SUBAPPLICATION AUF_AB_Softkey_Aux_DataPanel_QXA_SB (* Manuell Auf/Ab mit SoftKey+AUX auf DataPanel-MI-Ausgaenge, Anforderung Sperrblock *)
  (* Standard: 61499-2; Description: Copyright (c) 2026 Meisterschulen am Ostbahnhof This program and the accompanying materials are made available under the terms of the Eclipse Public License 2.0 which is available at https://www.eclipse.org/legal/epl-2.0/ SPDX-License-Identifier: EPL-2.0 *)
  (* Version 1.0, 2026-10-31, Franz Höpfinger, Meisterschulen am Ostbahnhof, Aus Getreidehacke func/Manual/ManFunc_AUF_AB3 in MyLib::sys verschoben und umbenannt, INIT/INITO/QI/QO ergaenzt, u8SAMember als Parameter. *)
  PACKAGE MyLib::sys;
  IMPORT isobus::UT::Q::const::IDs::ID_NULL;
  IMPORT DataPanel::io::MI::DQ::DataPanel_MI_DO_S;
  IMPORT DataPanel::io::MI::DQ::DataPanel_MI_DO;
  IMPORT DataPanel::io::MI::const::MI;
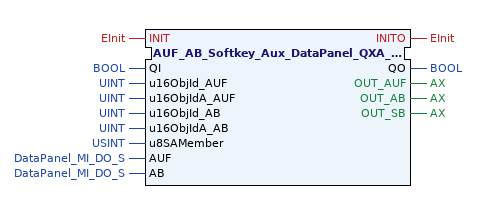
  EVENT_INPUT
    INIT : EInit; (* Initialization Request *)
  END_EVENT
  EVENT_OUTPUT
    INITO : EInit; (* Initialization Confirm *)
  END_EVENT
  VAR_INPUT
    QI : BOOL := TRUE; (* Quality Input - TRUE to enable service *)
    u16ObjId_AUF : UINT := ID_NULL; (* Object ID SoftKey AUF *)
    u16ObjIdA_AUF : UINT := ID_NULL; (* Object ID AuxFunction2 AUF *)
    u16ObjId_AB : UINT := ID_NULL; (* Object ID SoftKey AB *)
    u16ObjIdA_AB : UINT := ID_NULL; (* Object ID AuxFunction2 AB *)
    u8SAMember : USINT := MI::MI_00; (* DataPanel-MI-Modul (Source Address) *)
    AUF : DataPanel::io::MI::DQ::DataPanel_MI_DO_S := DataPanel_MI_DO::Invalid; (* DataPanel-MI-Ausgang AUF *)
    AB : DataPanel::io::MI::DQ::DataPanel_MI_DO_S := DataPanel_MI_DO::Invalid; (* DataPanel-MI-Ausgang AB *)
  END_VAR
  VAR_OUTPUT
    QO : BOOL; (* Quality Output - TRUE if service executed successfully *)
  END_VAR
  PLUGS
    OUT_AUF : adapter::types::unidirectional::AX; (* AUF aktiv *)
    OUT_AB : adapter::types::unidirectional::AX; (* AB aktiv *)
    OUT_SB : adapter::types::unidirectional::AX; (* Sperrblock anfordern (AUF ODER AB) *)
  END_PLUGS
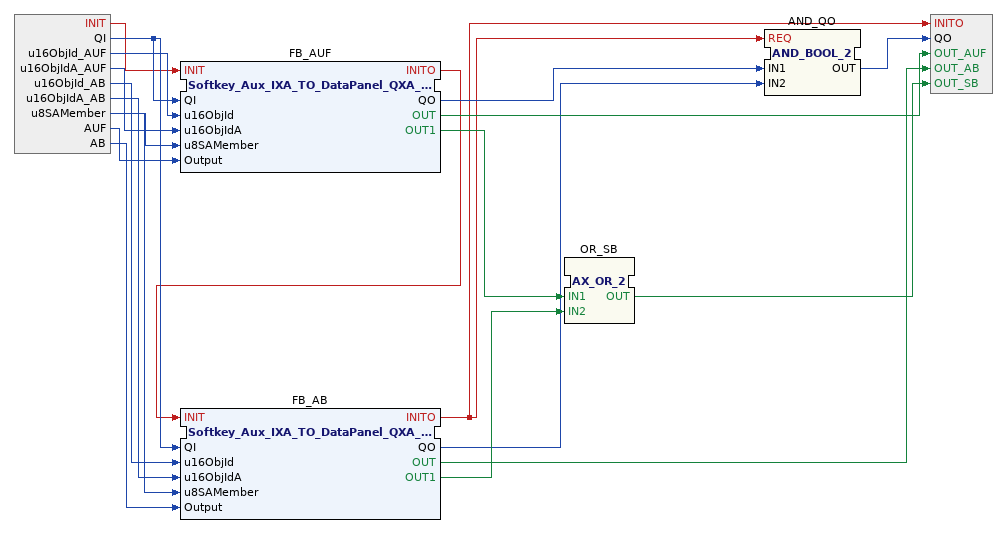
  FBS
    OR_SB : adapter::booleanOperators::AX_OR_2;
    AND_QO : iec61131::booleanOperators::AND_BOOL_2;
  END_FBS
  SUBAPPS
    FB_AUF : MyLib::sys::Softkey_Aux_IXA_TO_DataPanel_QXA_BG;
    FB_AB : MyLib::sys::Softkey_Aux_IXA_TO_DataPanel_QXA_BG;
  END_SUBAPPS
  EVENT_CONNECTIONS
    INIT TO FB_AUF.INIT;
    FB_AUF.INITO TO FB_AB.INIT;
    FB_AB.INITO TO INITO;
    FB_AB.INITO TO AND_QO.REQ;
  END_CONNECTIONS
  DATA_CONNECTIONS
    QI TO FB_AUF.QI;
    QI TO FB_AB.QI;
    u16ObjId_AUF TO FB_AUF.u16ObjId;
    u16ObjIdA_AUF TO FB_AUF.u16ObjIdA;
    u16ObjId_AB TO FB_AB.u16ObjId;
    u16ObjIdA_AB TO FB_AB.u16ObjIdA;
    u8SAMember TO FB_AUF.u8SAMember;
    u8SAMember TO FB_AB.u8SAMember;
    AUF TO FB_AUF.Output;
    AB TO FB_AB.Output;
    FB_AUF.QO TO AND_QO.IN1;
    FB_AB.QO TO AND_QO.IN2;
    AND_QO.OUT TO QO;
  END_CONNECTIONS
  ADAPTER_CONNECTIONS
    FB_AUF.OUT TO OUT_AUF;
    FB_AB.OUT TO OUT_AB;
    FB_AUF.OUT1 TO OR_SB.IN1;
    FB_AB.OUT1 TO OR_SB.IN2;
    OR_SB.OUT TO OUT_SB;
  END_CONNECTIONS
END_SUBAPPLICATION
